// TIA Portal V17 export
// export: Created 2026-11-08T05:50:29.4587933Z, ExportSetting WithDefaults, DisplayName Totally Integrated Automation Portal, DisplayVersion V17, DisplayName TIA Portal Openness, DisplayVersion V17, DisplayName TIA Portal Version Control Interface, DisplayVersion V17, DisplayName STEP 7 Professional, DisplayVersion V17, DisplayName STEP 7 Safety, DisplayVersion V17, DisplayName WinCC Professional, DisplayVersion V17
VAR_GLOBAL   // PLC tag table "Pilotos"
   HL_Marcha AT %M10.4 : Bool;   // Piloto verde: motor en marcha
   HL_Falla AT %M10.5 : Bool;   // Piloto rojo: falla térmico
END_VAR
